INTERFACE I_DifferentialDrive

METHOD Execute
END_METHOD

METHOD Enable
END_METHOD

METHOD Disable
END_METHOD

METHOD SetTwist
VAR_INPUT
	desiredTwist : Twist;
END_VAR
END_METHOD

PROPERTY LeftWheelPositionInM : LREAL
GET
END_GET
END_PROPERTY

PROPERTY RightWheelPositionInM : LREAL
GET
END_GET
END_PROPERTY

PROPERTY IsReady : BOOL
GET
END_GET
END_PROPERTY

END_INTERFACE

(* stored: Version 1.1.0.1, ProductVersion 3.1.4026.12
   Itf I_DifferentialDrive: Id {85909425-9268-52b7-9db9-1e67d6afd42c}
   Method Execute: Id {f5ce1296-efa5-51c7-a725-e150e3a9e895}
   Method Enable: Id {c017d325-fb79-52f8-9bdd-78a4ca5290c9}
   Method Disable: Id {e0109796-b129-527b-9f1e-df98fa7b3144}
   Method SetTwist: Id {117cb1ef-893c-5181-bcd7-b8426eef764c}
   Property LeftWheelPositionInM: Id {5e560f46-ced9-5ae6-a71f-0b50929bfbb4}
   Get Get: Id {e19dfd2b-29be-544f-9270-8290dd09801f}
   Property RightWheelPositionInM: Id {083f9cbc-56c2-56e7-999a-c7856fbac84b}
   Get Get: Id {e9258df9-3486-5059-ae42-043f5c11346e}
   Property IsReady: Id {1fff83d3-9da1-536a-a66d-02de1948d2fa}
   Get Get: Id {00c36e97-9830-5cca-886e-83179da3f416} *)
